Fanuc KAREL source: kb00198.KL

-- PROVISIONAL review KL for V940-1; original PC SHA256 fdc115d1c83e3ef8fc412958063fd01af777de67422e8d740b52b5247f990ac2
-- Incomplete behavior may be omitted. Consult companion uncertainty JSON. Do not deploy.
PROGRAM KB00198
%NOLOCKGROUP
BEGIN
  -- V9_ZERO_TABLE_METADATA_HINT layout=0002_ascii; no indexed target words; source/name/runtime held
  -- UNRESOLVED_PC offsets 5-14; opcodes 3F,75
  -- UNRESOLVED_PC offsets 19-26; opcodes 9D,23
  -- UNRESOLVED_PC offsets 31-38; opcodes 9D,23
  -- UNRESOLVED_PC offsets 43-79; opcodes 27,22,22,2A,22,22,22,31
  -- UNRESOLVED_PC offsets 84-88; opcodes 7F
END KB00198
